SUBAPPLICATION ILOCK_SWITCH_2_QXA_TASTER_OPC (* Kopie von ILOCK_SWITCH_2_QXA_OPC mit drittem Kommando-Eingang je Richtung (z.B. Hardware-Taster einer anderen Station, Remote-Subscribe) - Test, Funktion und Taster werden per AX_OR_3 zusammengefuehrt. Original: 2-Richtungs-Doppelwirkungs-Ausgang (Last-Wins mit Schutzzeit): je Richtung wird das echte Funktions-Kommando (Remote-Subscribe) mit dem bestehenden IO-Test-Kommando (Remote-Subscribe) per AX_OR_2 zusammengefuehrt, bevor es in den Interlock geht - IO-Test bleibt nutzbar, kann aber die beiden Richtungen nicht mehr dauerhaft gleichzeitig schalten. Interlocked Ausgang treibt den physischen logiBUS-Kanal UND meldet seinen tatsaechlichen Zustand sowohl an die bestehende IO-Test-Ueberwachung als auch an die echte Funktions-Rueckmeldung (z.B. GreenWhiteBackground am SoftKey) zurueck. Generisch fuer jeden 'digital DW'-Aktor (siehe IO-Liste_Vereinheitlicht.md) mit Bedienung von einem Modul ohne eigenes VT. *)
  (* Standard: 61499-2 *)
  (* Version 1.1, 2026-10-30, Franz Höpfinger, Meisterschulen am Ostbahnhof, INIT-Kette ohne Remote: SUBSCRIBE_TASTER_UP/DOWN (STG4 I4/I5, remote) nicht mehr seriell vor den Publishes, sondern parallel direkt an INIT, ohne Nachfolger. Damit entstehen Command/State-Nodes sofort mit der Option, auch wenn STG4 noch nicht da ist (sonst bis 60 s Remote-Init-Timeout, forte #1092). *)
  (* Version 1.0, 2026-10-17, Franz Höpfinger, Meisterschulen am Ostbahnhof, initial implementation - Kopie von ILOCK_SWITCH_2_QXA_OPC v1.3 (Original bleibt unveraendert), neue Eingaenge ID_TASTER_READ_UP/DOWN, OR_UP/OR_DOWN jetzt AX_OR_3, AND_QO jetzt AND_BOOL_12. Erstnutzung: Reihenverstellung KVE16 (Taster S1.7/S1.8 an STG4 I4/I5, Ventil an STG3 Q5/Q6). *)
  PACKAGE MyLib::sys;
  IMPORT logiBUS::io::DQ::logiBUS_DO;
  IMPORT logiBUS::io::DQ::logiBUS_DO_S;
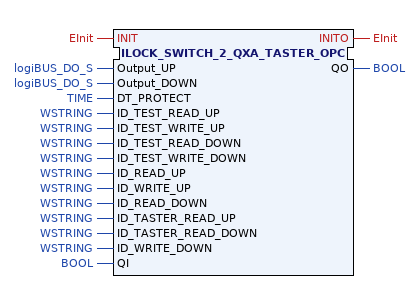
  EVENT_INPUT
    INIT : EInit; (* Initialisierung - vom Aufrufer sequenziert statt per Auto-Verteilung, damit QI vor der physischen Kanalbindung feststeht *)
  END_EVENT
  EVENT_OUTPUT
    INITO : EInit; (* Initialisierung bestaetigt (von DigitalOutput_UP.INITO) - fuer Aufrufer, die eine echte Confirm-Kette brauchen (z.B. hinter einem Option::AOption-Adapter) *)
  END_EVENT
  VAR_INPUT
    Output_UP : logiBUS::io::DQ::logiBUS_DO_S := logiBUS_DO::Invalid; (* Physischer Ausgang Richtung UP/Links *)
    Output_DOWN : logiBUS::io::DQ::logiBUS_DO_S := logiBUS_DO::Invalid; (* Physischer Ausgang Richtung DOWN/Rechts *)
    DT_PROTECT : TIME := T#300ms; (* Schutz-Totzeit vor Richtungswechsel *)
    ID_TEST_READ_UP : WSTRING; (* Bestehende IO-Test-Subscribe-Adresse UP (z.B. STG3_Q0x_READ) *)
    ID_TEST_WRITE_UP : WSTRING; (* Bestehende IO-Test-Publish-Adresse UP (z.B. STG3_Q0x_WRITE) *)
    ID_TEST_READ_DOWN : WSTRING; (* Bestehende IO-Test-Subscribe-Adresse DOWN *)
    ID_TEST_WRITE_DOWN : WSTRING; (* Bestehende IO-Test-Publish-Adresse DOWN *)
    ID_READ_UP : WSTRING; (* Echtes Funktions-Kommando UP (Subscribe) *)
    ID_WRITE_UP : WSTRING; (* Echte Funktions-Rueckmeldung UP (Publish) *)
    ID_READ_DOWN : WSTRING; (* Echtes Funktions-Kommando DOWN (Subscribe) *)
    ID_TASTER_READ_UP : WSTRING; (* Dritte Kommando-Quelle UP, z.B. Hardware-Taster (Subscribe) *)
    ID_TASTER_READ_DOWN : WSTRING; (* Dritte Kommando-Quelle DOWN, z.B. Hardware-Taster (Subscribe) *)
    ID_WRITE_DOWN : WSTRING; (* Echte Funktions-Rueckmeldung DOWN (Publish) *)
    QI : BOOL := TRUE; (* Qualifier fuer die physischen Ausgaenge - FALSE haelt diese Instanz komplett inaktiv (keine Hardware-Bindung), fuer den Fall dass derselbe physische Kanal je nach Maschinenvariante anderweitig genutzt wird *)
  END_VAR
  VAR_OUTPUT
    QO : BOOL; (* Quality Output - TRUE if service executed successfully (AND aller Subscribe/Publish/DigitalOutput-Instanzen) *)
  END_VAR
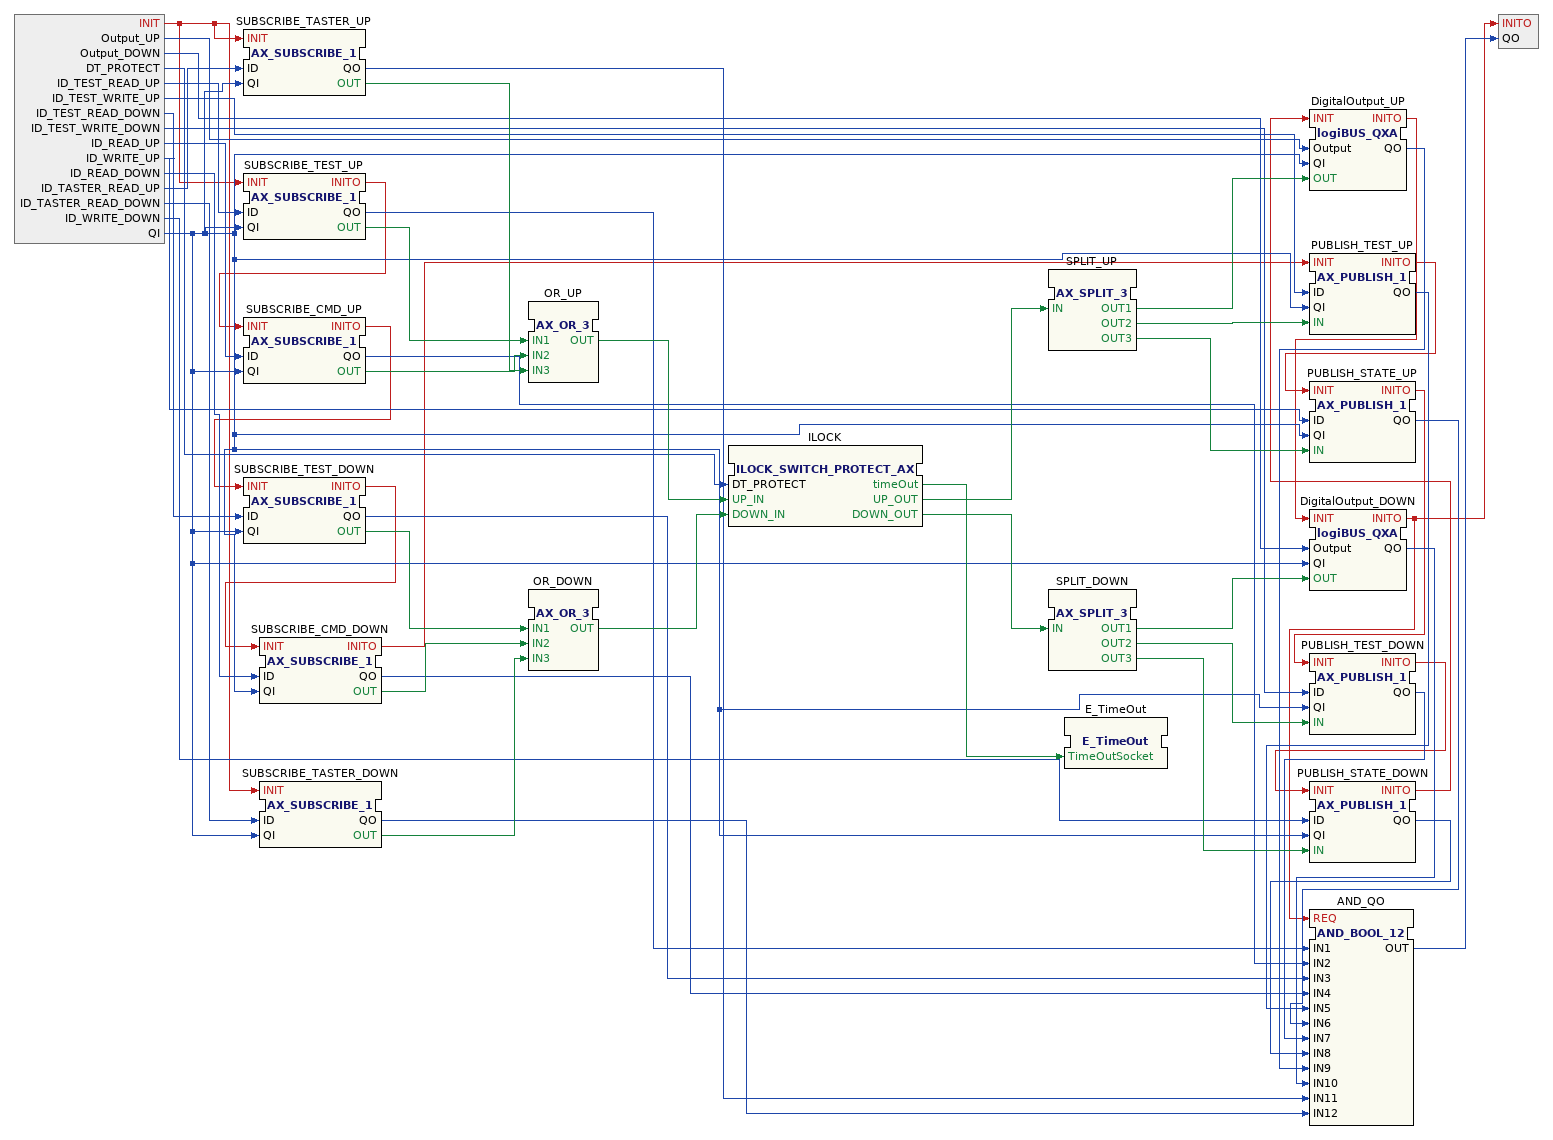
  FBS
    SUBSCRIBE_TEST_UP : adapter::net::AX_SUBSCRIBE_1;
    SUBSCRIBE_CMD_UP : adapter::net::AX_SUBSCRIBE_1;
    SUBSCRIBE_TASTER_UP : adapter::net::AX_SUBSCRIBE_1;
    SUBSCRIBE_TASTER_DOWN : adapter::net::AX_SUBSCRIBE_1;
    OR_UP : adapter::booleanOperators::AX_OR_3;
    SUBSCRIBE_TEST_DOWN : adapter::net::AX_SUBSCRIBE_1;
    SUBSCRIBE_CMD_DOWN : adapter::net::AX_SUBSCRIBE_1;
    OR_DOWN : adapter::booleanOperators::AX_OR_3;
    ILOCK : logiBUS::signalprocessing::interlock::ILOCK_SWITCH_PROTECT_AX;
    E_TimeOut : iec61499::events::E_TimeOut;
    SPLIT_UP : adapter::events::unidirectional::AX_SPLIT_3;
    SPLIT_DOWN : adapter::events::unidirectional::AX_SPLIT_3;
    DigitalOutput_UP : logiBUS::io::DQ::logiBUS_QXA;
    DigitalOutput_DOWN : logiBUS::io::DQ::logiBUS_QXA;
    PUBLISH_TEST_UP : adapter::net::AX_PUBLISH_1;
    PUBLISH_STATE_UP : adapter::net::AX_PUBLISH_1;
    PUBLISH_TEST_DOWN : adapter::net::AX_PUBLISH_1;
    PUBLISH_STATE_DOWN : adapter::net::AX_PUBLISH_1;
    AND_QO : iec61131::booleanOperators::AND_BOOL_12;
  END_FBS
  EVENT_CONNECTIONS
    INIT TO SUBSCRIBE_TEST_UP.INIT;
    SUBSCRIBE_TEST_UP.INITO TO SUBSCRIBE_CMD_UP.INIT;
    SUBSCRIBE_CMD_UP.INITO TO SUBSCRIBE_TEST_DOWN.INIT;
    SUBSCRIBE_TEST_DOWN.INITO TO SUBSCRIBE_CMD_DOWN.INIT;
    SUBSCRIBE_CMD_DOWN.INITO TO PUBLISH_TEST_UP.INIT;
    INIT TO SUBSCRIBE_TASTER_UP.INIT;
    INIT TO SUBSCRIBE_TASTER_DOWN.INIT;
    PUBLISH_TEST_UP.INITO TO PUBLISH_STATE_UP.INIT;
    PUBLISH_STATE_UP.INITO TO PUBLISH_TEST_DOWN.INIT;
    PUBLISH_TEST_DOWN.INITO TO PUBLISH_STATE_DOWN.INIT;
    PUBLISH_STATE_DOWN.INITO TO DigitalOutput_UP.INIT;
    DigitalOutput_UP.INITO TO DigitalOutput_DOWN.INIT;
    DigitalOutput_DOWN.INITO TO INITO;
    DigitalOutput_DOWN.INITO TO AND_QO.REQ;
  END_CONNECTIONS
  DATA_CONNECTIONS
    ID_TEST_READ_UP TO SUBSCRIBE_TEST_UP.ID;
    ID_READ_UP TO SUBSCRIBE_CMD_UP.ID;
    ID_TEST_READ_DOWN TO SUBSCRIBE_TEST_DOWN.ID;
    ID_READ_DOWN TO SUBSCRIBE_CMD_DOWN.ID;
    ID_TASTER_READ_UP TO SUBSCRIBE_TASTER_UP.ID;
    ID_TASTER_READ_DOWN TO SUBSCRIBE_TASTER_DOWN.ID;
    DT_PROTECT TO ILOCK.DT_PROTECT;
    Output_UP TO DigitalOutput_UP.Output;
    Output_DOWN TO DigitalOutput_DOWN.Output;
    QI TO DigitalOutput_UP.QI;
    QI TO DigitalOutput_DOWN.QI;
    ID_TEST_WRITE_UP TO PUBLISH_TEST_UP.ID;
    ID_WRITE_UP TO PUBLISH_STATE_UP.ID;
    ID_TEST_WRITE_DOWN TO PUBLISH_TEST_DOWN.ID;
    ID_WRITE_DOWN TO PUBLISH_STATE_DOWN.ID;
    QI TO SUBSCRIBE_TEST_UP.QI;
    QI TO SUBSCRIBE_CMD_UP.QI;
    QI TO SUBSCRIBE_TEST_DOWN.QI;
    QI TO SUBSCRIBE_CMD_DOWN.QI;
    QI TO SUBSCRIBE_TASTER_UP.QI;
    QI TO SUBSCRIBE_TASTER_DOWN.QI;
    QI TO PUBLISH_TEST_UP.QI;
    QI TO PUBLISH_STATE_UP.QI;
    QI TO PUBLISH_TEST_DOWN.QI;
    QI TO PUBLISH_STATE_DOWN.QI;
    SUBSCRIBE_TEST_UP.QO TO AND_QO.IN1;
    SUBSCRIBE_CMD_UP.QO TO AND_QO.IN2;
    SUBSCRIBE_TEST_DOWN.QO TO AND_QO.IN3;
    SUBSCRIBE_CMD_DOWN.QO TO AND_QO.IN4;
    PUBLISH_TEST_UP.QO TO AND_QO.IN5;
    PUBLISH_STATE_UP.QO TO AND_QO.IN6;
    PUBLISH_TEST_DOWN.QO TO AND_QO.IN7;
    PUBLISH_STATE_DOWN.QO TO AND_QO.IN8;
    DigitalOutput_UP.QO TO AND_QO.IN9;
    DigitalOutput_DOWN.QO TO AND_QO.IN10;
    SUBSCRIBE_TASTER_UP.QO TO AND_QO.IN11;
    SUBSCRIBE_TASTER_DOWN.QO TO AND_QO.IN12;
    AND_QO.OUT TO QO;
  END_CONNECTIONS
  ADAPTER_CONNECTIONS
    SUBSCRIBE_TEST_UP.OUT TO OR_UP.IN1;
    SUBSCRIBE_CMD_UP.OUT TO OR_UP.IN2;
    SUBSCRIBE_TASTER_UP.OUT TO OR_UP.IN3;
    OR_UP.OUT TO ILOCK.UP_IN;
    SUBSCRIBE_TEST_DOWN.OUT TO OR_DOWN.IN1;
    SUBSCRIBE_CMD_DOWN.OUT TO OR_DOWN.IN2;
    SUBSCRIBE_TASTER_DOWN.OUT TO OR_DOWN.IN3;
    OR_DOWN.OUT TO ILOCK.DOWN_IN;
    ILOCK.timeOut TO E_TimeOut.TimeOutSocket;
    ILOCK.UP_OUT TO SPLIT_UP.IN;
    SPLIT_UP.OUT1 TO DigitalOutput_UP.OUT;
    SPLIT_UP.OUT2 TO PUBLISH_TEST_UP.IN;
    SPLIT_UP.OUT3 TO PUBLISH_STATE_UP.IN;
    ILOCK.DOWN_OUT TO SPLIT_DOWN.IN;
    SPLIT_DOWN.OUT1 TO DigitalOutput_DOWN.OUT;
    SPLIT_DOWN.OUT2 TO PUBLISH_TEST_DOWN.IN;
    SPLIT_DOWN.OUT3 TO PUBLISH_STATE_DOWN.IN;
  END_CONNECTIONS
END_SUBAPPLICATION
